		//481 -----------------------------------
		,(code		:= 17198
		,message 	:= '17198.  DWORD for the interpretation of the axis units not allowed The value that contains the flags for the interpretation of the position and velocity units is not allowed.')
		//482 -----------------------------------
		,(code		:= 17199
		,message 	:= '17199.  Maximum velocity not allowed The value for the maximum permitted velocity is not allowed.')
		//483 -----------------------------------
		,(code		:= 17200
		,message 	:= '17200.  Motion monitoring window not allowed The value for the motion monitoring window is not allowed. V')
		//484 -----------------------------------
		,(code		:= 17201
		,message 	:= '17201.  PEH time monitoring not allowed The value for the activation of the PEH time monitoring is not allowed (PEH: positioning end and halt).')
		//485 -----------------------------------
		,(code		:= 17202
		,message 	:= '17202.  PEH monitoring time not allowed The value for the PEH monitoring time (timeout) is not allowed (PEH: positioning end and halt). Default value: 5 s')
		//486 -----------------------------------
		,(code		:= 17203
		,message 	:= '17203.  AXISERR_RANGE_DELAYBREAKRELEASE')
		//487 -----------------------------------
		,(code		:= 17204
		,message 	:= '17204.  ?AXISERR_RANGE_DATAPERSISTENCE?')
		//488 -----------------------------------
		,(code		:= 17210
		,message 	:= '17210.  ?AXISERR_RANGE_POSDIFF_FADING_ACCELERATION?')
		//489 -----------------------------------
		,(code		:= 17211
		,message 	:= '17211.  Fast Axis Stop Signal Type not allowed The value for the Signal Type of the Fast Axis Stop is not allowed [0...5].')
		//490 -----------------------------------
		,(code		:= 17216
		,message 	:= '17216.  Axis initialisation Axis has not been initialised. Although the axis has been created, the rest of the initialisation has not been performed (1. Initialisation of axis I/O, 2. Initialisation of axis, 3. Reset axis).')
		//491 -----------------------------------
		,(code		:= 17217
		,message 	:= '17217.  Group address Axis does not have a group, or the group address has not been initialised (group contains the set value generation).')
		//492 -----------------------------------
		,(code		:= 17218
		,message 	:= '17218.  Encoder address The axis does not have an encoder, or the encoder address has not been initialised.')
		//493 -----------------------------------
		,(code		:= 17219
		,message 	:= '17219.  Controller address The axis does not have a controller, or the controller address has not been initialised.')
		//494 -----------------------------------
		,(code		:= 17220
		,message 	:= '17220.  Drive address The axis does not have a drive, or the drive address has not been initialised.')
		//495 -----------------------------------
		,(code		:= 17221
		,message 	:= '17221.  Axis interface PLC to NC address Axis does not have an axis interface from the PLC to the NC, or the axis interface address has not been initialised.')
		//496 -----------------------------------
		,(code		:= 17222
		,message 	:= '17222.  Axis interface NC to PLC address Axis does not have an axis interface from the NC to the PLC, or the axis interface address has not been initialised.')
		//497 -----------------------------------
		,(code		:= 17223
		,message 	:= '17223.  Size of axis interface NC to PLC is not allowed (INTERNAL ERROR) The size of the axis interface from NC to PLC is not allowed.')
		//498 -----------------------------------
		,(code		:= 17224
		,message 	:= '17224.  Size of axis interface PLC to NC is not allowed (INTERNAL ERROR) The size of the axis interface from PLC to NC is not allowed.')
		//499 -----------------------------------
		,(code		:= 17238
		,message 	:= '17238.  Controller enable Controller enable for the axis is not present (see axis interface SPS®NC). This enable is required, for instance, for an axis positioning task.')
		//500 -----------------------------------
		,(code		:= 17239
		,message 	:= '17239.  Feed enable minus Feed enable for movement in the negative direction is not present (see axis interface SPS®NC). This enable is required, for instance, for an axis positioning task in the negative direction.')
		//501 -----------------------------------
		,(code		:= 17240
		,message 	:= '17240.  Feed enable plus Feed enable for movement in the positive direction is not present (see axis interface SPS®NC). This enable is required, for instance, for an axis positioning task in the positive direction.')
		//502 -----------------------------------
		,(code		:= 17241
		,message 	:= '17241.  Set velocity not allowed The set velocity requested for a positioning task is not allowed. This can happen if the velocity is less than or equal to zero, larger than the maximum permitted axis velocity, or, in the case of servo-drives, is larger than the reference velocity of the axis (see axis and drive parameters).')
		//503 -----------------------------------
		,(code		:= 17242
		,message 	:= '17242.  Movement smaller than one encoder increment (INTERNAL ERROR) The movement required of an axis is, in relation to a positioning task, smaller than one encoder increment (see scaling factor). This information is, however, handled internally in such a way that the positioning is considered to have been completed without an error message being returned.')
		//504 -----------------------------------
		,(code		:= 17243
		,message 	:= '17243.  Set acceleration monitoring (INTERNAL ERROR) The set acceleration has exceeded the maximum permitted acceleration or deceleration parameters of the axis.')
		//505 -----------------------------------
		,(code		:= 17244
		,message 	:= '17244.  PEH time monitoring The PEH time monitoring has detected that, after the PEH monitoring time that follows a positioning has elapsed, the target position window has not been reached. The following points must be checked: Is the PEH monitoring time, in the sense of timeout monitoring, set to a sufficiently large value (e.g. 1-5s)? The PEH monitoring time must be chosen to be significantly larger than the target position monitoring time. Have the criteria for the target position monitoring (range window and time) been set too strictly?')
		//506 -----------------------------------
		,(code		:= 17245
		,message 	:= '17245.  Encoder existence monitoring / movement monitoring During the active positioning the actual encoder value has changed continuously for a default check time from NC cycle to NC cycle less than the default minimum movement limit.')
		//507 -----------------------------------
		,(code		:= 17246
		,message 	:= '17246.  ?Looping distance less than breaking distance? The absolute value of the looping distance is less or equal than the positive or negative breaking distance. This is not allowed.')
		//508 -----------------------------------
		,(code		:= 17249
		,message 	:= '17249.  ?Time range exceeded (future)? The calculated position lies too far in the future (e.g. when converting a position value in a DC time stamp).')
		//509 -----------------------------------
		,(code		:= 17250
		,message 	:= '17250.  ?Time range exceeded (past)? The calculated position lies too far in the past (e.g. when converting a position value in a DC time stamp).')
		//510 -----------------------------------
		,(code		:= 17251
		,message 	:= '17251.  ?Position cannot be determined? The requested position cannot be determined.')
		//511 -----------------------------------
		,(code		:= 17312
		,message 	:= '17312.  Axis consequential error Consequential error resulting from another causative error related to another axis. Axis consequential errors can occur in relation to master/slave couplings or with multiple axis interpolating DXD groups.')
		//512 -----------------------------------
		,(code		:= 17408
		,message 	:= '17408.  Encoder ID not allowed The value for the encoder ID is not allowed, e.g. because it has already been assigned, is less than or equal to zero, or is bigger than 255.')
		//513 -----------------------------------
		,(code		:= 17409
		,message 	:= '17409.  Encoder type not allowed The value for the encoder type is unacceptable because it is not defined. Type 1: Simulation (incremental) Type 2: M3000 (24 bit absolute) Type 3: M31x0 (24 bit incremental) Type 4: KL5101 (16 bit incremental) Type 5: KL5001 (24 bit absolute SSI) Type 6: KL5051 (16 bit BISSI)')
		//514 -----------------------------------
		,(code		:= 17410
		,message 	:= '17410.  Encoder mode The value for the encoder (operating) mode is not allowed. Mode 1: Determination of the actual position Mode 2: Determination of the actual position and the actual velocity (filter)')
		//515 -----------------------------------
		,(code		:= 17411
		,message 	:= '17411.  Encoder counting direction inverted? The flag for the encoder counting direction is not allowed. Flag 0: Positive encoder counting direction Flag 1: Negative encoder counting direction')
		//516 -----------------------------------
		,(code		:= 17412
		,message 	:= '17412.  Referencing status The flag for the referencing status is not allowed. Flag 0: Axis has not been referenced Flag 1: Axis has been referenced')
		//517 -----------------------------------
		,(code		:= 17413
		,message 	:= '17413.  Encoder increments for each physical encoder rotation The value for the number of encoder increments for each physical rotation of the encoder is not allowed. This value is used by the software for the calculation of encoder overruns and underruns.')
		//518 -----------------------------------
		,(code		:= 17414
		,message 	:= '17414.  Scaling factor The value for the scaling factor is not allowed. This scaling factor provides the weighting for the conversion of an encoder increment (INC) to a physical unit such as millimeters or degrees.')
		//519 -----------------------------------
		,(code		:= 17415
		,message 	:= '17415.  Position offset (zero point offset) The value for the position offset of the encoder is not allowed. This value is added to the calculated encoder position, and is interpreted in the physical units of the encoder.')
		//520 -----------------------------------
		,(code		:= 17416
		,message 	:= '17416.  Modulo factor The value for the encoders modulo factor is not allowed.')
		//521 -----------------------------------
		,(code		:= 17417
		,message 	:= '17417.  Position filter time The value for the actual position filter time is not allowed (P-T1 filter).')
		//522 -----------------------------------
		,(code		:= 17418
		,message 	:= '17418.  Velocity filter time The value for the actual velocity filter time is not allowed (P-T1 filter).')
		//523 -----------------------------------
		,(code		:= 17419
		,message 	:= '17419.  Acceleration filter time The value for the actual acceleration filter time is not allowed (P-T1 filter).')
		//524 -----------------------------------
		,(code		:= 17420
		,message 	:= '17420.  Cycle time not allowed (INTERNAL ERROR) The value of the SAF cycle time for the calculation of actual values is not allowed (e.g. is less than or equal to zero).')
		//525 -----------------------------------
		,(code		:= 17421
		,message 	:= '17421.  ENCERR_RANGE_UNITFLAGS')
		//526 -----------------------------------
		,(code		:= 17422
		,message 	:= '17422.  Actual position correction / measurement system error correction The value for the activation of the actual position correction (measuring system error correction) is not allowed.')
		//527 -----------------------------------
		,(code		:= 17423
		,message 	:= '17423.  Filter time actual position correction The value for the actual position correction filter time is not allowed (P-T1 filter).')
		//528 -----------------------------------
		,(code		:= 17424
		,message 	:= '17424.  Search direction for referencing cam inverted The value of the search direction of the referencing cam in a referencing procedure is not allowed. Value 0: Positive direction Value 1: Negative direction')
		//529 -----------------------------------
		,(code		:= 17425
		,message 	:= '17425.  Search direction for sync pulse (zero pulse) inverted The value of the search direction of the sync pulse (zero pulse) in a referencing procedure is not allowed. Value 0: Positive direction Value 1: Negative direction')
		//530 -----------------------------------
		,(code		:= 17426
		,message 	:= '17426.  Reference position The value of the reference position in a referencing procedure is not allowed.')
		//531 -----------------------------------
		,(code		:= 17427
		,message 	:= '17427.  Clearance monitoring between activation of the hardware latch and appearance of the sync pulse (NOT IMPLEMENTED) The flag for the clearance monitoring between activation of the hardware latch and occurrence of the sync/zero pulse (latch valid) is not allowed. Value 0: Passive Value 1: Active')
		//532 -----------------------------------
		,(code		:= 17428
		,message 	:= '17428.  Minimum clearance between activation of the hardware latch and appearance of the sync pulse (NOT IMPLEMENTED) The value for the minimum clearance in increments between activation of the hardware latch and occurrence of the sync/zero pulse (latch valid) during a referencing procedure is not allowed.')
		//533 -----------------------------------
		,(code		:= 17429
		,message 	:= '17429.  External sync pulse (NOT IMPLEMENTED) The value of the activation or deactivation of the external sync pulse in a referencing procedure is not allowed. Value 0: Passive Value 1: Active')
		//534 -----------------------------------
		,(code		:= 17430
		,message 	:= '17430.  Scaling of the noise rate is not allowed The value of the scaling (weighting) of the synthetic noise rate is not allowed. This parameter exists only in the simulation encoder and serves to produce a realistic simulation.')
		//535 -----------------------------------
		,(code		:= 17431
		,message 	:= '17431.  ?Tolerance window for modulo-start? The value for the tolerance window for the modulo-axis-start is invalid. The value must be greater or equal than zero and smaller than the half encoder modulo-period (e. g. in the interval [0.0,180.0) ).')
		//536 -----------------------------------
		,(code		:= 17432
		,message 	:= '17432.  ?Encoder reference mode? The value for the encoder reference mode is not allowed, resp. is not supported for this encoder type.')
		//537 -----------------------------------
		,(code		:= 17433
		,message 	:= '17433.  ?Encoder evaluation direction? The value for the encoder evaluation direction (log. counter direction) is not allowed.')
		//538 -----------------------------------
		,(code		:= 17434
		,message 	:= '17434.  ?Encoder reference system? The value for the encoder reference system is invalid (0: incremental, 1: absolute, 2: absolute+modulo).')
		//539 -----------------------------------
		,(code		:= 17435
		,message 	:= '17435.  ?Encoder position initialization mode? When starting the TC system the value for the encoder position initialization mode is invalid.')
		//540 -----------------------------------
		,(code		:= 17436
		,message 	:= '17436.  ?Encoder sign interpretation (UNSIGNED- / SIGNED- data type)? The value for the encoder sign interpretation (data type) for the encoder the actual increment calculation (0: Default/not defined, 1: UNSIGNED, 2:/ SIGNED) is invalid.')
		//541 -----------------------------------
		,(code		:= 17440
		,message 	:= '17440.  Software end location monitoring minimum not allowed The value for the activation of the software location monitoring minimum is not allowed.')
		//542 -----------------------------------
		,(code		:= 17441
		,message 	:= '17441.  Software end location monitoring maximum not allowed The value for the activation of the software location monitoring maximum is not allowed.')
		//543 -----------------------------------
		,(code		:= 17442
		,message 	:= '17442.  Actual value setting is outside the value range The set actual value function cannot be carried out, because the new actual position is outside the expected range of values.')
		//544 -----------------------------------
		,(code		:= 17443
		,message 	:= '17443.  Software end location minimum not allowed The value for the software end location minimum is not allowed.')
		//545 -----------------------------------
		,(code		:= 17444
		,message 	:= '17444.  Software end location maximum not allowed The value for the software end location maximum is not allowed.')
		//546 -----------------------------------
		,(code		:= 17445
		,message 	:= '17445.  ?Filter mask for the raw data of the encoder is invalid? The value for the filter mask of the encoder raw data in increments is invalid.')
		//547 -----------------------------------
		,(code		:= 17446
		,message 	:= '17446.  ?Reference mask for the raw data of the encoder is invalid? The value for the reference mask (increments per encoder turn, absolute resolution) for the raw data of the encoder is invalid. E.g. this value is used for axis reference sequence (calibration) with the reference mode Software Sync.')
		//548 -----------------------------------
		,(code		:= 17456
		,message 	:= '17456.  Hardware latch activation (encoder) Activation of the encoder hardware latch was implicitly initiated by the referencing procedure. If this function has already been activated but a latch value has not yet become valid (latch valid), another call to the function is refused with this error.')
		//549 -----------------------------------
		,(code		:= 17457
		,message 	:= '17457.  External hardware latch activation (encoder) The activation of the external hardware latch (only available on the KL5101) is initiated explicitly by an ADS command (called from the PLC program of the Visual Basic interface). If this function has already been activated, but the latch value has not yet been made valid by an external signal (external latch valid), another call to the function is refused with this error.')
		//550 -----------------------------------
		,(code		:= 17458
		,message 	:= '17458.  External hardware latch activation (encoder) If a referencing procedure has previously been initiated and the hardware still signals a valid latch value (latch valid), this function must not be called. In practice, however, this error can almost never occur.')
		//551 -----------------------------------
		,(code		:= 17459
		,message 	:= '17459.  External hardware latch activation (encoder) If this function has already been initiated and the hardware is still signaling that the external latch value is still valid (extern latch valid), a further activation should not be carried out and the commando will be declined with an error (the internal handshake communication between NC and IO device is still active). In that case the validity of the external hardware latch would immediately be signaled, although the old latch value would still be present.')
		//552 -----------------------------------
		,(code		:= 17460
		,message 	:= '17460.  Encoder function not supported An encoder function has been activated that is currently not released for use, or which is not even implemented.')
		//553 -----------------------------------
		,(code		:= 17461
		,message 	:= '17461.  ?Encoder function is already active? An encoder function can not been activated because this functionality is already active.')
		//554 -----------------------------------
		,(code		:= 17472
		,message 	:= '17472.  Encoder initialization Encoder has not been initialized. Although the axis has been created, the rest of the initialization has not been performed (1. Initialization of axis I/O, 2. Initialization of axis, 3. Reset axis).')
		//555 -----------------------------------
		,(code		:= 17473
		,message 	:= '17473.  Axis address The encoder does not have an axis, or the axis address has not been initialized.')
		//556 -----------------------------------
		,(code		:= 17474
		,message 	:= '17474.  I/O input structure address The drive does not have a valid I/O input address in the process image.')
		//557 -----------------------------------
		,(code		:= 17475
		,message 	:= '17475.  I/O output structure address The encoder does not have a valid I/O output address in the process image.')
		//558 -----------------------------------
		,(code		:= 17488
		,message 	:= '17488.  Encoder counter underflow monitoring The encoders incremental counter has underflowed.')
		//559 -----------------------------------
		,(code		:= 17489
		,message 	:= '17489.  Encoder counter overflow monitoring The encoders incremental counter has overflowed.')
		//560 -----------------------------------
		,(code		:= 17504
		,message 	:= '17504.  Software end location minimum (axis start) With active monitoring of the software end location for a minimum, a start has been made from a position that lies below the software end location minimum.')
		//561 -----------------------------------
		,(code		:= 17505
		,message 	:= '17505.  Software end location maximum (axis start) With active monitoring of the software end location for a maximum, a start has been made from a position that lies above the software end location maximum.')
		//562 -----------------------------------
		,(code		:= 17506
		,message 	:= '17506.  Software end location minimum (positioning process) With active monitoring of the software end location for a minimum, the actual position has fallen below the software end location minimum. In the case of servo axes (continuously driven axes) this limit is expanded by the magnitude of the parameterized following error window (position).')
		//563 -----------------------------------
		,(code		:= 17507
		,message 	:= '17507.  Software end location maximum (positioning process) With active monitoring of the software end location for a maximum, the actual position has exceeded the software end location maximum. In the case of servo axes (continuously driven axes) this limit is expanded by the magnitude of the parameterized following error window (position).')
		//564 -----------------------------------
		,(code		:= 17508
		,message 	:= '17508.  ?Encoder hardware error? The drive resp. the encoder system reports a hardware error of the encoder. An optimal error code is displayed in the message of the event log.')
		//565 -----------------------------------
		,(code		:= 17509
		,message 	:= '17509.  ?Position initialization error at system start? At the first initialization of the set position was this for all initialization trials (without over-/under-flow, with underflow and overflow ) out of the final position minimum and maximum.')
		//566 -----------------------------------
		,(code		:= 17520
		,message 	:= '17520.  SSI transformation fault or not finished The SSI transformation of the FOX 50 module was faulty for some NC-cycles or did not finished respectively.')
		//567 -----------------------------------
		,(code		:= 17570
		,message 	:= '17570.  ENCERR_ADDR_CONTROLLER')
		//568 -----------------------------------
		,(code		:= 17571
		,message 	:= '17571.  ENCERR_INVALID_CONTROLLERTYPE')
		//569 -----------------------------------
		,(code		:= 17664
		,message 	:= '17664.  Controller ID not allowed The value for the controller ID is not allowed, e.g. because it has already been assigned, is less than or equal to zero, or is greater than 255.')
		//570 -----------------------------------
		,(code		:= 17665
		,message 	:= '17665.  Controller type not allowed The value for the controller type is unacceptable because it is not defined. Type 1: P-controller (position) . . . Type 7: High/low speed controller Type 8: Stepper motor controller Type 9: Sercos controller')
		//571 -----------------------------------
		,(code		:= 17666
		,message 	:= '17666.  Controller operating mode not allowed The value for the controller operating mode is not allowed.')
		//572 -----------------------------------
		,(code		:= 17667
		,message 	:= '17667.  Weighting of the velocity pre-control not allowed The value for the percentage weighting of the velocity pre-control is not allowed. The parameter is pre-set to 1.0 (100%) as standard.')
		//573 -----------------------------------
		,(code		:= 17668
		,message 	:= '17668.  Following error monitoring (position) not allowed The value for the activation of the following error monitoring is not allowed.')
		//574 -----------------------------------
		,(code		:= 17669
		,message 	:= '17669.  Following error (velocity) not allowed The value for the activation of the following error monitoring (velocity) is not allowed.')
		//575 -----------------------------------
		,(code		:= 17670
		,message 	:= '17670.  Following error window (position) not allowed The value for the following error window (maximum allowable following error) is not allowed.')
		//576 -----------------------------------
		,(code		:= 17671
		,message 	:= '17671.  Following error filter time (position) not allowed The value for the following error filter time (position) is not allowed.')
		//577 -----------------------------------
		,(code		:= 17672
		,message 	:= '17672.  Following error window (velocity) not allowed The value for the following error window (velocity) is not allowed.')
		//578 -----------------------------------
		,(code		:= 17673
		,message 	:= '17673.  Following error filter time (velocity) not allowed The value for the following error filter time (velocity) is not allowed.')
		//579 -----------------------------------
		,(code		:= 17680
		,message 	:= '17680.  Proportional gain Kv or Kp (position controller) not allowed The value for the proportional gain (Kv factor or Kp factor) is not allowed.')
		//580 -----------------------------------
		,(code		:= 17681
		,message 	:= '17681.  Integral-action time Tn (position controller) not allowed The value for the integral-action time is not allowed (I proportion of the PID T1 controller).')
		//581 -----------------------------------
		,(code		:= 17682
		,message 	:= '17682.  Derivative action time Tv (position controller) not allowed The value for the derivative action time is not allowed (D proportion of the PID T1 controller).')
		//582 -----------------------------------
		,(code		:= 17683
		,message 	:= '17683.  Damping time Td (position controller) not allowed The value for the damping time is not allowed (D proportion of the PID T1 controller). Suggested value: 0.1 * Tv')
		//583 -----------------------------------
		,(code		:= 17684
		,message 	:= '17684.  Activation of the automatic offset compensation not allowed Activation of the automatic offset compensation is only possible for certain types of controller (with no I component).')
		//584 -----------------------------------
		,(code		:= 17685
		,message 	:= '17685.  Additional proportional gain Kv or Kp (position controller) not allowed The value for the second term of the proportional gain (Kv factor or Kp factor) is not allowed.')
		//585 -----------------------------------
		,(code		:= 17686
		,message 	:= '17686.  Reference velocity for additional proportional gain Kv or Kp (positioncontroller) not allowed The value for the reference velocity percentage data entry, to which the additional proportional gain is applied, is not allowed. The standard setting for the parameter is 0.5 (50%).')
		//586 -----------------------------------
		,(code		:= 17687
		,message 	:= '17687.  Proportional gain Pa (acceleration proportion) not allowed The value for the proportional gain (Pa factor) is not allowed.')
		//587 -----------------------------------
		,(code		:= 17688
		,message 	:= '17688.  Proportional gain Kv (velocity controller) not allowed The value for the proportional gain (Kv factor) is not allowed.')
		//588 -----------------------------------
		,(code		:= 17689
		,message 	:= '17689.  ?Reset time Tn (velocity controller) not allowed? The value for the integral-action time is not allowed (I proportion of the PID T1 controller).')
		//589 -----------------------------------
		,(code		:= 17690
		,message 	:= '17690.  CONTROLERR_RANGE_ACCJUMPLIMITINGMODE')
		//590 -----------------------------------
		,(code		:= 17691
		,message 	:= '17691.  CONTROLERR_RANGE_ACCJUMPVALUE')
		//591 -----------------------------------
		,(code		:= 17692
		,message 	:= '17692.  CONTROLERR_RANGE_FILTERTIME')
		//592 -----------------------------------
		,(code		:= 17693
		,message 	:= '17693.  ?Dead zone not allowed? The value for the dead zone from the position error or the velocity error (system deviation) is not allowed (only for complex controller with velocity or torque interface).')
		//593 -----------------------------------
		,(code		:= 17696
		,message 	:= '17696.  ?Rate time Tv (velocity controller) not allowed? The value for the derivative action time is not allowed (D proportion of the PID T1 controller).')
		//594 -----------------------------------
		,(code		:= 17697
		,message 	:= '17697.  Damping time Td (velocity controller) not allowed The value for the damping time is not allowed (D proportion of the PID T1 controller). Suggested value: 0.1 * Tv')
		//595 -----------------------------------
		,(code		:= 17698
		,message 	:= '17698.  CONTROLERR_RANGE_IOUTPUTLIMIT')
		//596 -----------------------------------
		,(code		:= 17699
		,message 	:= '17699.  CONTROLERR_RANGE_DOUTPUTLIMIT')
		//597 -----------------------------------
		,(code		:= 17700
		,message 	:= '17700.  CONTROLERR_RANGE_POSIDISABLEWHENMOVING')
		//598 -----------------------------------
		,(code		:= 17728
		,message 	:= '17728.  Controller initialisation Controller has not been initialised. Although the controller has been created, the rest of the initialisation has not been performed (1. Initialisation of controller, 2. Reset controller).')
		//599 -----------------------------------
		,(code		:= 17729
		,message 	:= '17729.  Axis address Controller does not know its axis, or the axis address has not been initialised.')
		//600 -----------------------------------
		,(code		:= 17730
		,message 	:= '17730.  Drive address Controller does not know its drive, or the drive address has not been initialised.')
		//601 -----------------------------------
		,(code		:= 17744
		,message 	:= '17744.  Following error monitoring (position) With active following error monitoring (position) a following error exceedance has occurred, whose magnitude is greater than the following error window, and whose duration is longer than the parameterised following error filter time.')
		//602 -----------------------------------
		,(code		:= 17745
		,message 	:= '17745.  Following error monitoring (velocity) With active following error monitoring (velocity) a velocity following error exceedance has occurred, whose magnitude is greater than the following error window, and whose duration is longer than the parameterised following error filter time.')
		//603 -----------------------------------
		,(code		:= 17824
		,message 	:= '17824.  CONTROLERR_RANGE_AREA_ASIDE')
		//604 -----------------------------------
		,(code		:= 17825
		,message 	:= '17825.  CONTROLERR_RANGE_AREA_BSIDE')
		//605 -----------------------------------
		,(code		:= 17826
		,message 	:= '17826.  CONTROLERR_RANGE_QNENN')
		//606 -----------------------------------
		,(code		:= 17827
		,message 	:= '17827.  CONTROLERR_RANGE_PNENN')
		//607 -----------------------------------
		,(code		:= 17828
		,message 	:= '17828.  CONTROLERR_RANGE_AXISIDPRESP0')
		//608 -----------------------------------
		,(code		:= 17920
		,message 	:= '17920.  Drive ID not allowed The value for the drive ID is not allowed, e.g. because it has already been assigned, is less than or equal to zero, or is greater than 255.')
		//609 -----------------------------------
		,(code		:= 17921
		,message 	:= '17921.  Drive type not allowed The value for the drive type is unacceptable because it is not defined.')
		//610 -----------------------------------
		,(code		:= 17922
		,message 	:= '17922.  Drive operating mode not allowed The value for the drive operating mode is not allowed. Modus 1:       Standard')
		//611 -----------------------------------
		,(code		:= 17923
		,message 	:= '17923.  Motor polarity inverted? The flag for the motor polarity is not allowed. Flag 0: Positive motor polarity Flag 1: Negative motor polarity')
		//612 -----------------------------------
		,(code		:= 17924
		,message 	:= '17924.  Drift compensation/velocity offset (DAC offset) The value for the drift compensation (DAC offset) is not allowed.')
		//613 -----------------------------------
		,(code		:= 17925
		,message 	:= '17925.  Reference velocity (velocity pre-control) The value for the reference velocity (velocity pre-control) is not allowed.')
		//614 -----------------------------------
		,(code		:= 17926
		,message 	:= '17926.  Reference output in percent The value for the reference output in percent is not allowed. The value 1.0 (100 %) usually corresponds to a voltage of 10.0 V.')
		//615 -----------------------------------
		,(code		:= 17927
		,message 	:= '17927.  Quadrant compensation factor The value for the quadrant compensation factor is not allowed.')
		//616 -----------------------------------
		,(code		:= 17928
		,message 	:= '17928.  Velocity reference point in percent The value for the velocity reference point in percent is not allowed. The value 1.0 corresponds to 100 percent.')
		//617 -----------------------------------
		,(code		:= 17929
		,message 	:= '17929.  Output reference point in percent The value for the output reference point in percent is not allowed. The value 1.0 corresponds to 100 percent.')
		//618 -----------------------------------
		,(code		:= 17930
		,message 	:= '17930.  Minimum or maximum output limit The values for the minimum and/or maximum output limit is not allowed. This will happen if the range of values is exceeded, the maximum limit is smaller than the minimum limit, or the distance between the minimum and maximum limits is zero. The minimum limit is initially set to 1.0 (-100 percent) and the maximum limit to 1.0 (100 percent).')
		//619 -----------------------------------
		,(code		:= 17931
		,message 	:= '17931.  DRIVEERR_RANGE_MAXINCREMENT')
		//620 -----------------------------------
		,(code		:= 17932
		,message 	:= '17932.  DRIVEERR_RANGE_ DRIVECONTROLDWORD')
		//621 -----------------------------------
		,(code		:= 17933
		,message 	:= '17933.  DRIVEERR_RANGE_ RESETCYCLECOUNTER')
		//622 -----------------------------------
		,(code		:= 17935
		,message 	:= '17935.  ?Drive torque output scaling is not allowed? The value for the drive torque output scaling (rotary motor) or the force output scaling (linear motor) is not allowed.')
		//623 -----------------------------------
		,(code		:= 17936
		,message 	:= '17936.  ?Drive velocity output scaling is not allowed? The value for the drive velocity output scaling is not allowed.')
		//624 -----------------------------------
		,(code		:= 17937
		,message 	:= '17937.  Profi Drive DSC Proportional gain  Kpc (position controller) not allowed The value for the profi drive DSC proportional gain (Kpc factor) is not allowed.')
		//625 -----------------------------------
		,(code		:= 17938
		,message 	:= '17938.  ?Table-ID is invalid? The value for the table-ID is invalid.')
		//626 -----------------------------------
		,(code		:= 17939
		,message 	:= '17939.  ?Table interpolationtype is invalid? The value for the table interpolation-type is invalid.')
		//627 -----------------------------------
		,(code		:= 17940
		,message 	:= '17940.  ?Outputoffset in percent is invalid? The value for the output offset in percent (+/- 1.0) is invalid.')
		//628 -----------------------------------
		,(code		:= 17941
		,message 	:= '17941.  ?Profi Drive DSC scaling factor for calculating Xerr (position controller) is not allowed? The value as profi drive DSC scaling factor for calculating Xerr is invalid.')
		//629 -----------------------------------
		,(code		:= 17942
		,message 	:= '17942.  ?Drive acceleration output scaling is not allowed? The value for the drive acceleration/deceleration output scaling is not allowed.')
		//630 -----------------------------------
		,(code		:= 17943
		,message 	:= '17943.  ?Drive position output scaling is not allowed? The value for the drive position output scaling is not allowed.')
		//631 -----------------------------------
		,(code		:= 17948
		,message 	:= '17948.  ?Drive filter typ for reference position variable is not allowed? The value for the drive filter type of the reference position output filter is not allowed.')
		//632 -----------------------------------
		,(code		:= 17949
		,message 	:= '17949.  ?Drive filter time for reference position variable is not allowed? The value for the drive filter time of the reference position output filter is not allowed.')
		//633 -----------------------------------
		,(code		:= 17950
		,message 	:= '17950.  ?Drive filter order for reference position variable is not allowed? The value for the drive filter order (P-Tn) of the reference position output filter is not allowed.')
		//634 -----------------------------------
		,(code		:= 17952
		,message 	:= '17952.  Bit mask for stepper motor cycle not allowed A value in the various stepper motor masks for the cycle concerned is not allowed.')
		//635 -----------------------------------
		,(code		:= 17953
		,message 	:= '17953.  Bit mask for stepper motor holding current not allowed The value for the stepper motor holding mask is not allowed.')
		//636 -----------------------------------
		,(code		:= 17968
		,message 	:= '17968.  ?Overtemperature? The drive resp. terminal detects an overtemperature alarm.')
		//637 -----------------------------------
		,(code		:= 17969
		,message 	:= '17969.  ?Undervoltage? The drive resp. terminal detects an undervoltage (supply voltage to low).')
		//638 -----------------------------------
		,(code		:= 17970
		,message 	:= '17970.  ?Wire breakage in phase A? The drive resp. terminal detects a wire breakage in phase A.')
		//639 -----------------------------------
		,(code		:= 17971
		,message 	:= '17971.  ?Wire breakage in phase B? The drive resp. terminal detects a wire breakage in phase B.')
		//640 -----------------------------------
		,(code		:= 17972
		,message 	:= '17972.  ?Overcurrent in phase A? The drive resp. terminal detects an overcurrent in phase A.')
		//641 -----------------------------------
		,(code		:= 17973
		,message 	:= '17973.  ?Overcurrent in Phase B? The drive resp. terminal detects an overcurrent in phase B.')
		//642 -----------------------------------
		,(code		:= 17974
		,message 	:= '17974.  ?Torque overload (stall situation)? The drive resp. terminal detects a torque overload (stall situation).')
		//643 -----------------------------------
		,(code		:= 17984
		,message 	:= '17984.  Drive initialisation Drive has not been initialised. Although the drive has been created, the rest of the initialisation has not been performed (1. Initialisation of drive I/O, 2. Initialisation of drive, 3. Reset drive).')
		//644 -----------------------------------
		,(code		:= 17985
		,message 	:= '17985.  Axis address Drive does not know its axis, or the axis address has not been initialised.')
		//645 -----------------------------------
		,(code		:= 17986
		,message 	:= '17986.  I/O input structure address The drive does not have a valid I/O input address in the process image.')
		//646 -----------------------------------
		,(code		:= 17987
		,message 	:= '17987.  I/O output structure address The drive does not have a valid I/O output address in the process image.')
		//647 -----------------------------------
		,(code		:= 18000
		,message 	:= '18000.  Drive not ready for operation The drive is not ready for operation. The following are possible causes: - the drive is in failure state (hardware fault) - the drive is in the starting-up stage (e.g. following an axis reset preceded by a hardware fault) - the drive has not been enabled Remark: The time required for booting a drive after a hardware fault can amount to several seconds.')
		//648 -----------------------------------
		,(code		:= 18001
		,message 	:= '18001.  Error in cyclic communication with the drive (life counter)')
		//649 -----------------------------------
		,(code		:= 18002
		,message 	:= '18002.  Not permitted to change the table ID while the axis is enabled')
		//650 -----------------------------------
		,(code		:= 18005
		,message 	:= '18005.  Invalid IO data for more than n consecutive nc cycles')
		//651 -----------------------------------
		,(code		:= 18944
		,message 	:= '18944.  Table ID not allowed The value for the table ID is not allowed, e.g. because it has already been assigned, is less than or equal to zero, or is greater than 255.')
		//652 -----------------------------------
		,(code		:= 18945
		,message 	:= '18945.  Table type not allowed The value for the table type is unacceptable because it is not defined.')
		//653 -----------------------------------
		,(code		:= 18946
		,message 	:= '18946.  Number of lines in the table not allowed The value of the number of lines in the table is not allowed, because, for example, it is smaller than two at linear interpolation and smaller than four at spline interpolation.')
		//654 -----------------------------------
		,(code		:= 18947
		,message 	:= '18947.  Number of columns in the table is not allowed The value of the number of columns in the table is not allowed, because, for example, it is less than or equal to zero (depends upon the type of table or slave).')
		//655 -----------------------------------
		,(code		:= 18948
		,message 	:= '18948.  Step size (position delta) not allowed The value for the step size between two lines (position delta) is not allowed, because, for example, it is less than or equal to zero.')
		//656 -----------------------------------
		,(code		:= 18949
		,message 	:= '18949.  Period not allowed The value for the period is not allowed, because, for example, it is less than or equal to zero.')
		//657 -----------------------------------
		,(code		:= 18950
		,message 	:= '18950.  Table is not monotonic The value for the step size is not allowed, because, for example, it is less than or equal to zero.')
		//658 -----------------------------------
		,(code		:= 18951
		,message 	:= '18951.  ?Table sub type is not allowed? The value for the table sub type is not allowed or otherwise the table class (slave type) do not match up to the table main type.')
		//659 -----------------------------------
		,(code		:= 18952
		,message 	:= '18952.  ?Table interpolation type is not allowed? The value for the table interpolation type is allowed.')
		//660 -----------------------------------
		,(code		:= 18953
		,message 	:= '18953.  Incorrect table main type The table main type is unknown or otherwise the table class (slave type) do not match up to the table main type.')
		//661 -----------------------------------
		,(code		:= 18960
		,message 	:= '18960.  Table initialisation Table has not been initialised. Although the table has been created, the rest of the initialisation has not been performed. For instance, the number of lines or columns may be less than or equal to zero.')
		//662 -----------------------------------
		,(code		:= 18961
		,message 	:= '18961.  Not enough memory Table could not be created, since there is not enough memory.')
		//663 -----------------------------------
		,(code		:= 18962
		,message 	:= '18962.  Function not executed, function not available The function has not been implemented, or cannot be executed, for the present type of table.')
		//664 -----------------------------------
		,(code		:= 18963
		,message 	:= '18963.  Line index not allowed The start line index or the stop line index to be used for read or write access to the table is not allowed. For instance, the line index may be greater than the total number of lines in the table.')
		//665 -----------------------------------
		,(code		:= 18964
		,message 	:= '18964.  Column index not allowed The start column index or the stop column index to be used for read or write access to the table in not allowed. For instance, the column index may be greater than the total number of columns in the table.')
		//666 -----------------------------------
		,(code		:= 18965
		,message 	:= '18965.  Number of lines not allowed The number of lines to be read from or written to the table is not allowed. The number of lines must be an integer multiple of the number of elements in a line (n * number of columns).')
		//667 -----------------------------------
		,(code		:= 18966
		,message 	:= '18966.  Number of columns not allowed The number of columns to be read from or written to the table is not allowed. The number of columns must be an integer multiple of the number of elements in a column (n * number of lines).')
		//668 -----------------------------------
		,(code		:= 18967
		,message 	:= '18967.  Error in scaling or in range entry The entries in the table header are inconsistent, e.g. the validity range is empty. If the error is generated during the run time it is a run time error and stops the master/slave group.')
		//669 -----------------------------------
		,(code		:= 18968
		,message 	:= '18968.  Multi table slave out of range The slave master position is outside the table values for the master. The error is a run-time error, and stops the master/slave group.')
		//670 -----------------------------------
		,(code		:= 18969
		,message 	:= '18969.  Solo table underflow The slave master position is outside the table values for the master. The master value of the equidistant table, to be processed linearly, lies under the first table value. The error is a run-time error, and stops the master/slave group.')
		//671 -----------------------------------
		,(code		:= 18970
		,message 	:= '18970.  Solo table overflow The slave master position is outside the table values for the master. The master value of the equidistant table, to be processed linearly, lies above the first table value. The error is a run-time error, and stops the master/slave group.')
		//672 -----------------------------------
		,(code		:= 18971
		,message 	:= '18971.  Incorrect execution mode The cyclic execution mode can only be true or false.')
		//673 -----------------------------------
		,(code		:= 18972
		,message 	:= '18972.  Impermissible parameter The Fifo parameter is not allowed.')
		//674 -----------------------------------
		,(code		:= 18973
		,message 	:= '18973.  Fifo is empty The Fifo of the external generator is empty. This can signify end of track or a run time error.')
		//675 -----------------------------------
		,(code		:= 18974
		,message 	:= '18974.  Fifo is full The Fifo of the external generator is full. It is the user?s task to continue to attempt to fill the Fifo with the rejected values.')
		//676 -----------------------------------
		,(code		:= 18975
		,message 	:= '18975.  ?Point-Index of Motion Function invalid?  The point index of a Motion Function Point of a Function Table is invalid. First the point index has to be larger than zero and second it has to be numerical continuously for one column in the Montion Function Table (e.g. 1,2,3,... or 10,11,12,...).')
		//677 -----------------------------------
		,(code		:= 18976
		,message 	:= '18976.  ?No diagonalisation of  matrix? The spline can not be calculated. The master positions are not correct.')
		//678 -----------------------------------
		,(code		:= 18977
		,message 	:= '18977.  ?Number of spline points to less? The number of points of a cubic spline has to be greater than two.')
		//679 -----------------------------------
		,(code		:= 18978
		,message 	:= '18978.  ?Fifo must not be overwritten? Fifo must not be overwritten since then the active line would be overwritten. It is the task of the user to secure that the active line is not modified.')
		//680 -----------------------------------
		,(code		:= 18979
		,message 	:= '18979.  ?Insufficient number of Motion Function points? The number of valid Motion Function points is less than two. Either the entire number of points is to low or the point type of many points is set to Ignore Point.')
		//681 -----------------------------------
		,(code		:= 19200
		,message 	:= '19200.  Axis has been stopped The axis has been stopped while the axis moves to target position. The axis could be stopped with a PLC Command via ADS, with the call of AXFNC or with the TwinCAT System Manager.')
		//682 -----------------------------------
		,(code		:= 19201
		,message 	:= '19201.  Axis cannot be started The axis cannot be started, because:')
		//683 -----------------------------------
		,(code		:= 19202
		,message 	:= '19202.  Control mode not allowed No Target Position Control and no Position Area Control.')
		//684 -----------------------------------
		,(code		:= 19203
		,message 	:= '19203.  Axis is not moving Restart position and velocity is only allowed if axis is physically moving.')
		//685 -----------------------------------
		,(code		:= 19204
		,message 	:= '19204.  Wrong mode for RestartPosAndVelo Wrong mode.')
		//686 -----------------------------------
		,(code		:= 19205
		,message 	:= '19205.  Command not allowed')
		//687 -----------------------------------
		,(code		:= 19206
		,message 	:= '19206.  Parameter not correct')
		//688 -----------------------------------
		,(code		:= 19207
		,message 	:= '19207.  Timeout axis function block Exact position cannot be reached with active current limit, but is not far enough off to cause following error.')
		//689 -----------------------------------
		,(code		:= 19208
		,message 	:= '19208.  Axis in protected mode Axis is in protected mode (i.e. coupled) and cannot be moved.')
		//690 -----------------------------------
		,(code		:= 19209
		,message 	:= '19209.  Axis is not ready Axis is not ready and cannot be moved.')
		//691 -----------------------------------
		,(code		:= 19210
		,message 	:= '19210.  Homing error The Homing of an axis could not be started or was not successful')
		//692 -----------------------------------
		,(code		:= 19211
		,message 	:= '19211.  Invalid definition trigger input definition The definition of the trigger signal used with the function block MC_TouchProbe is invalid. The defined encoder ID, the trigger signal or the trigger signal edge are invalid.')
		//693 -----------------------------------
		,(code		:= 19212
		,message 	:= '19212.  position latch has been deactivated The function block MC_TouchProbe encountered that a touch probe sequence has been deactivated after the block started this sequence. The reason for instance can be an axis reset.')
		//694 -----------------------------------
		,(code		:= 19213
		,message 	:= '19213.  Timeout NC status feedback A function block has successfully executed a command but the NC does not pass the expected feedback in the axis status word.')
		//695 -----------------------------------
		,(code		:= 19214
		,message 	:= '19214.  Supplement not installed - The function is available as supplement product but not installed on the system.')
		//696 -----------------------------------
		,(code		:= 19215
		,message 	:= '19215.  Timeout Register Access - The access to a bus terminal register timed out.')
		//697 -----------------------------------
		,(code		:= 19216
		,message 	:= '19216.  M-Function request missing This error occurs if a confirmation of an M-Function is made but the request bit is not set.')
		//698 -----------------------------------
		,(code		:= 19217
		,message 	:= '19217.  Zero shift index is out of range The index of the zero shift is invalid')
		//699 -----------------------------------
		,(code		:= 19218
		,message 	:= '19218.  R parameter index or size is invalid. This error occurs, if the R parameters are written or read and the index or size is out of range')
		//700 -----------------------------------
		,(code		:= 19219
		,message 	:= '19219.  Index for tool description is invalid')
		//701 -----------------------------------
		,(code		:= 19220
		,message 	:= '19220.  Version of cyclic channel interface does not match to the requested function and function block, resp. This error occurs, if an older TwinCAT Version is used and a new functionality from a newer TcNci.lib is called.')
		//702 -----------------------------------
		,(code		:= 19221
		,message 	:= '19221.  Channel is not ready for requested function. The requested function can not be executed due to a wrong state of the channel. This error occurs for instance, if retrace is requested and the axes are not stopped with ItpEStop before.')
		//703 -----------------------------------
		,(code		:= 19222
		,message 	:= '19222.  Requested function is not turned on. The requested function requires an explicit activation before it can be executed.')
		//704 -----------------------------------
		,(code		:= 19232
		,message 	:= '19232.  Cannot append all axes. This error occurs, if you want to append an auxiliary axes to an interpolation group and the function fails. Probably a prior assignment of an auxiliary axes was skipped.')
		//705 -----------------------------------
		,(code		:= 19248
		,message 	:= '19248.  Pointer invalid. The pointer to a data structure is invalid, e.g. NULL.')
		//706 -----------------------------------
		,(code		:= 19249
		,message 	:= '19249.  Size of  memory invalid. The size parameter is invalid.')
		//707 -----------------------------------
		,(code		:= 19250
		,message 	:= '19250.  Invalid cam table ID. The cam table ID is out of the range from 1 to 255.')
		//708 -----------------------------------
		,(code		:= 19251
		,message 	:= '19251.  Invalid point ID. The point ID of a motion function point is lower than 1.')
		//709 -----------------------------------
		,(code		:= 19252
		,message 	:= '19252.  Invalid number of points . The number of points to read or write is less than 1.')
		//710 -----------------------------------
		,(code		:= 19253
		,message 	:= '19253.  Invalid MC table type. The type of a cam table does not match theMC_TableType definition.')
		//711 -----------------------------------
		,(code		:= 19254
		,message 	:= '19254.  Invalid number of rows. The number of rows of a cam table is less than 1.')
		//712 -----------------------------------
		,(code		:= 19255
		,message 	:= '19255.  Invalid number of columns. The number of columns of a cam table is invalid.')
		//713 -----------------------------------
		,(code		:= 19256
		,message 	:= '19256.  Invalid Increment. The increment for an interpolation is invalid, e.g. <= 0.')
		//714 -----------------------------------
		,(code		:= 19264
		,message 	:= '19264.  Unsupported Terminal Type.  The terminal in use is not supported by this function block.')
		//715 -----------------------------------
		,(code		:= 19265
		,message 	:= '19265.  Register Read/Write Error.   This error implies to be a validation error.')
		//716 -----------------------------------
		,(code		:= 19266
		,message 	:= '19266.  Axis is Enabled.  Axis is enabled and is not supposed to be enabled for this operation')
		//717 -----------------------------------
		,(code		:= 19267
		,message 	:= '19267.  Size of compensation table wrong. The stated table size in bytes is not conform with the real size.')
		//718 -----------------------------------
		,(code		:= 19268
		,message 	:= '19268.  The minimum/ maximum position of the compenstation table is not conform to the position in the table description (ST_CompensationDesc)')
		//719 -----------------------------------
		,(code		:= 19269
		,message 	:= '19269.  Not implemented. The requested function is not implemented in this combination.')
		//720 -----------------------------------
		,(code		:= 19296
		,message 	:= '19296.  Motion command not be activated. A motion command has been started and has been buffered and confirmed by the NC. Nevertheless the command did not become active.')
		//721 -----------------------------------
		,(code		:= 19297
		,message 	:= '19297.  Motion command could not be monitored by the PLC. A motion command has been started and has been buffered and confirmed by the NC. The PLC has not been able to monitor the execution of this command and the execution status is unclear since the NC is already executing a more recent command. This error may com up with very short buffered motion commands which are executed during one PLC cycle.')
		//722 -----------------------------------
		,(code		:= 19298
		,message 	:= '19298.  Buffered command finished with error. A buffered command finished with an error. The error number is not available because a new command is already in execution.')
		//723 -----------------------------------
		,(code		:= 19299
		,message 	:= '19299.  Buffered command finished without state feedback. A buffered command finished without success or error feedback.')
		//724 -----------------------------------
		,(code		:= 19300
		,message 	:= '19300.  BufferMode not supported. The BufferMode is not supported by the command.')
		//725 -----------------------------------
		,(code		:= 19301
		,message 	:= '19301.  Command number is zero. The system administrated command number for buffered commands is zero.')
		//726 -----------------------------------
		,(code		:= 19302
		,message 	:= '19302.  Function block was not called cyclically . The function block was not called cyclically and the PLC was therefore not able to monitor the motion command while the NC is already executing another command. The execution state is unclear.')
		//727 -----------------------------------
		,(code		:= 19313
		,message 	:= '19313.  Invalid NCI Entry Type. FB_NciFeedTablePreparation is called with an unknown nEntryType')
		//728 -----------------------------------
		,(code		:= 19314
		,message 	:= '19314.  NciFeedTable full. The table is full filled and therefore this entry is not accepted.')
		//729 -----------------------------------
		,(code		:= 19315
		,message 	:= '19315.  internal error')
		//730 -----------------------------------
		,(code		:= 19316
		,message 	:= '19316.  ST_NciTangentialFollowingDesc: tangential axis is not an auxiliary axis The entry ST_NciTangentialFollowingDesc contains an tangential axis that is no auxiliary axis.')
		//731 -----------------------------------
		,(code		:= 19317
		,message 	:= '19317.  ST_NciTangentialFollowingDesc: nPathAxis1 and nPathAxis2, resp. are no path axes. So it is not possible to determine the plane.')
		//732 -----------------------------------
		,(code		:= 19318
		,message 	:= '19318.  ST_NciTangentialFollwoingDesc: nPathAxis1 and nPathAxis2 are equal. So it is not possible to determine the plane.')
		//733 -----------------------------------
		,(code		:= 19319
		,message 	:= '19319.  ST_NciGeoCirclePlane: circle is programmed in a wrong manner.')
		//734 -----------------------------------
		,(code		:= 19320
		,message 	:= '19320.  Internal error in calculation of the tangential following')
		//735 -----------------------------------
		,(code		:= 19321
		,message 	:= '19321.  Tangential following: With ST_NciTangentialFollowingDesc the monitoring of the deviation angle (E_TfErrorOnCrirical1) is activated and with the actual segment the deviation angle is too big.')
		//736 -----------------------------------
		,(code		:= 19322
		,message 	:= '19322.  not implemented')
		//737 -----------------------------------
		,(code		:= 19323
		,message 	:= '19323.  Tangential Following: The radius of the actual circle segment is too small')
		//738 -----------------------------------
		,(code		:= 19324
		,message 	:= '19324.  FB_NciFeedTablePreparation:  pEntry is NULL')
		//739 -----------------------------------
		,(code		:= 19325
		,message 	:= '19325.  FB_NciFeedTablePreparation: The specified nEntryType does not match the the structure type')
		//740 -----------------------------------
		,(code		:= 19326
		,message 	:= '19326.  ST_NciMFuncFast and ST_NciMFuncHsk: The requested m-function is not in between 0..159')
		//741 -----------------------------------
		,(code		:= 19327
		,message 	:= '19327.  ST_NciDynOvr: The requested value for the dynamic override is not in between 0.01 and 1.0')
		//742 -----------------------------------
		,(code		:= 19328
		,message 	:= '19328.  ST_NciVertexSmoothing: invalid parameter. This error occurs with a negative vertex radius or an unknown vertex smoothing type.')
		//743 -----------------------------------
		,(code		:= 19329
		,message 	:= '19329.  FB_NciFeedTablePrepartion: The requested velocity is not in a valid range')
		//744 -----------------------------------
		,(code		:= 19330
		,message 	:= '19330.  ST_Nci*: invalid parameter')
	]
	;
	{warning restore C0198}
END_VAR

(* stored: Version 1.1.0.1, ProductVersion 3.1.4024.12
   GVL GVL_Lib_TcErrors: Id {bfc89e73-e3b6-47df-9fd7-08f67411cd19} *)
